(* IEC 61131-3 sources: kns-pump-station/tests/POUs/Station/FB_PumpRotation_Test, 30 files *)

(* ---- AdoptAtPlcStartFromFeedback.method.decl.st ---- *)
// 04 §13.3, PMI-35: старт ПЛК — подхват по ОС (GVL_IO.xP10n_RFB) до первого вызова устройства; запрос не снимается
// ни недоступностью первого цикла, ни ограничением последовательного пуска
METHOD PRIVATE AdoptAtPlcStartFromFeedback
VAR
    fbDut    : FB_PumpRotation;                    // ФБ под тестом
    fbTime   : PL.FB_FakeTime;                     // подменное время, старт 1 ч
    stCfg    : ST_StationCfg;                      // уставки по умолчанию (RunHours, tStagger 5 с)
    stRetain : ST_StationRetain;                   // следующий ведущий (Cyclic)
    afbPump  : ARRAY[1..3] OF FB_FakeMotorVfd;     // подменные насосы: доступны, Auto, готовы, стоят
    fbSink   : FB_FakeEventSink;                   // подменный журнал
END_VAR

(* ---- AdoptKeepsRunningPumpsOnAutoEntry.method.decl.st ---- *)
// 04 §3.2, PMI-30: вход в «Автомат» — роли получают работающие насосы (ещё в Manual в этом цикле), работающий не
// останавливается, ведущий — с меньшей наработкой
METHOD PRIVATE AdoptKeepsRunningPumpsOnAutoEntry
VAR
    fbDut    : FB_PumpRotation;                    // ФБ под тестом
    fbTime   : PL.FB_FakeTime;                     // подменное время, старт 1 ч
    stCfg    : ST_StationCfg;                      // уставки по умолчанию (RunHours, tStagger 5 с)
    stRetain : ST_StationRetain;                   // следующий ведущий (Cyclic)
    afbPump  : ARRAY[1..3] OF FB_FakeMotorVfd;     // подменные насосы: доступны, Auto, готовы, стоят
    fbSink   : FB_FakeEventSink;                   // подменный журнал
END_VAR

(* ---- Cycle.method.decl.st ---- *)
// Помощник: uiSteps шагов времени tStep с одним требуемым числом. xPlant — подменные насосы в Auto
// следуют запросам: работают, если запрошены, доступны и без отказа (видно со следующего шага)
METHOD PRIVATE Cycle
VAR_IN_OUT
    fbDut    : FB_PumpRotation;                 // ФБ под тестом
    fbTime   : PL.FB_FakeTime;                  // подменное время
    stCfg    : ST_StationCfg;                   // уставки
    stRetain : ST_StationRetain;                // энергонезависимые данные
    afbPump  : ARRAY[1..3] OF FB_FakeMotorVfd;  // подменные насосы
END_VAR
VAR_INPUT
    uiRequired : UINT;                          // требуемое число насосов
    tStep      : TIME;                          // шаг времени
    uiSteps    : UINT;                          // шагов
    xPlant     : BOOL;                          // насосы следуют запросам
END_VAR
VAR
    uiStep : UINT;                              // номер шага
    uiIdx  : UINT;                              // насос
END_VAR

(* ---- Cycle.method.impl.st ---- *)
FOR uiStep := 1 TO uiSteps DO
    fbTime.Advance(tStep := tStep);
    fbDut(uiRequired := uiRequired, itfTime := fbTime, stCfg := stCfg, stRetain := stRetain);
    IF xPlant THEN
        FOR uiIdx := 1 TO 3 DO
            IF afbPump[uiIdx].eMode = PL.E_DeviceMode.Auto THEN
                afbPump[uiIdx].xRunning := fbDut.axRun[uiIdx] AND afbPump[uiIdx].xAvailable
                                           AND NOT afbPump[uiIdx].xFault;
            END_IF
        END_FOR
    END_IF
END_FOR

(* ---- CyclicAdvancesNextLeadRetained.method.decl.st ---- *)
// 04 §8.1, PMI-10: по кругу — ведущий после stStationRetain.uiNextLead независимо от наработки, следующий
// запоминается энергонезависимо
METHOD PRIVATE CyclicAdvancesNextLeadRetained
VAR
    fbDut    : FB_PumpRotation;                    // ФБ под тестом
    fbTime   : PL.FB_FakeTime;                     // подменное время, старт 1 ч
    stCfg    : ST_StationCfg;                      // уставки по умолчанию (RunHours, tStagger 5 с)
    stRetain : ST_StationRetain;                   // следующий ведущий (Cyclic)
    afbPump  : ARRAY[1..3] OF FB_FakeMotorVfd;     // подменные насосы: доступны, Auto, готовы, стоят
    fbSink   : FB_FakeEventSink;                   // подменный журнал
END_VAR

(* ---- CyclicNextLeadFollowsRoleTransfer.method.decl.st ---- *)
// 04 §8.1, §8.2, PMI-10, PMI-11: по кругу следующий ведущий отсчитывается от насоса, который стал ведущим, в том
// числе без нового пуска (передача роли по ограничению непрерывной работы). Иначе после передачи Н1 → Н2
// следующий пуск снова достался бы Н2, а Н3 простаивал бы
METHOD PRIVATE CyclicNextLeadFollowsRoleTransfer
VAR
    fbDut    : FB_PumpRotation;                    // ФБ под тестом
    fbTime   : PL.FB_FakeTime;                     // подменное время, старт 1 ч
    stCfg    : ST_StationCfg;                      // уставки по умолчанию, режим Cyclic
    stRetain : ST_StationRetain;                   // следующий ведущий (Cyclic)
    afbPump  : ARRAY[1..3] OF FB_FakeMotorVfd;     // подменные насосы: доступны, Auto, готовы, стоят
    fbSink   : FB_FakeEventSink;                   // подменный журнал
END_VAR

(* ---- CyclicStopsAssist.method.decl.st ---- *)
// 04 §5.2: по кругу и без чередования — при уменьшении останавливается подпорный
METHOD PRIVATE CyclicStopsAssist
VAR
    fbDut    : FB_PumpRotation;                    // ФБ под тестом
    fbTime   : PL.FB_FakeTime;                     // подменное время, старт 1 ч
    stCfg    : ST_StationCfg;                      // уставки по умолчанию (RunHours, tStagger 5 с)
    stRetain : ST_StationRetain;                   // следующий ведущий (Cyclic)
    afbPump  : ARRAY[1..3] OF FB_FakeMotorVfd;     // подменные насосы: доступны, Auto, готовы, стоят
    fbSink   : FB_FakeEventSink;                   // подменный журнал
END_VAR

(* ---- DisabledNoRequestsRolesStandby.method.decl.st ---- *)
// DESIGN 6.5: станция не в «Автомате» — запросов нет, роли считаются (Standby у доступных, None у недоступных)
METHOD PRIVATE DisabledNoRequestsRolesStandby
VAR
    fbDut    : FB_PumpRotation;                    // ФБ под тестом
    fbTime   : PL.FB_FakeTime;                     // подменное время, старт 1 ч
    stCfg    : ST_StationCfg;                      // уставки по умолчанию (RunHours, tStagger 5 с)
    stRetain : ST_StationRetain;                   // следующий ведущий (Cyclic)
    afbPump  : ARRAY[1..3] OF FB_FakeMotorVfd;     // подменные насосы: доступны, Auto, готовы, стоят
    fbSink   : FB_FakeEventSink;                   // подменный журнал
END_VAR

(* ---- EmergencyRequiresAllThree.method.decl.st ---- *)
// 04 §10.2, PMI-20: аварийный режим — запросы всем трём насосам по одному через tStagger; роли Lead, Assist,
// Assist
METHOD PRIVATE EmergencyRequiresAllThree
VAR
    fbDut    : FB_PumpRotation;                    // ФБ под тестом
    fbTime   : PL.FB_FakeTime;                     // подменное время, старт 1 ч
    stCfg    : ST_StationCfg;                      // уставки по умолчанию (RunHours, tStagger 5 с)
    stRetain : ST_StationRetain;                   // следующий ведущий (Cyclic)
    afbPump  : ARRAY[1..3] OF FB_FakeMotorVfd;     // подменные насосы: доступны, Auto, готовы, стоят
    fbSink   : FB_FakeEventSink;                   // подменный журнал
END_VAR

(* ---- FaultedPumpLosesRequestImmediately.method.decl.st ---- *)
// 04 §9.1, PMI-12, PMI-13: отказавший ведущий теряет запрос сразу (роль None), замена — в том же вызове
METHOD PRIVATE FaultedPumpLosesRequestImmediately
VAR
    fbDut    : FB_PumpRotation;                    // ФБ под тестом
    fbTime   : PL.FB_FakeTime;                     // подменное время, старт 1 ч
    stCfg    : ST_StationCfg;                      // уставки по умолчанию (RunHours, tStagger 5 с)
    stRetain : ST_StationRetain;                   // следующий ведущий (Cyclic)
    afbPump  : ARRAY[1..3] OF FB_FakeMotorVfd;     // подменные насосы: доступны, Auto, готовы, стоят
    fbSink   : FB_FakeEventSink;                   // подменный журнал
END_VAR

(* ---- FixedOrder.method.decl.st ---- *)
// 04 §8.1: без чередования — Н1, Н2, Н3 по порядку; недоступный пропускается
METHOD PRIVATE FixedOrder
VAR
    fbDut    : FB_PumpRotation;                    // ФБ под тестом
    fbTime   : PL.FB_FakeTime;                     // подменное время, старт 1 ч
    stCfg    : ST_StationCfg;                      // уставки по умолчанию (RunHours, tStagger 5 с)
    stRetain : ST_StationRetain;                   // следующий ведущий (Cyclic)
    afbPump  : ARRAY[1..3] OF FB_FakeMotorVfd;     // подменные насосы: доступны, Auto, готовы, стоят
    fbSink   : FB_FakeEventSink;                   // подменный журнал
END_VAR

(* ---- ForeignRunningReducesRequests.method.decl.st ---- *)
// 04 §5.1, PMI-31: сторонний работающий насос (не в Auto) уменьшает число запросов станции
METHOD PRIVATE ForeignRunningReducesRequests
VAR
    fbDut    : FB_PumpRotation;                    // ФБ под тестом
    fbTime   : PL.FB_FakeTime;                     // подменное время, старт 1 ч
    stCfg    : ST_StationCfg;                      // уставки по умолчанию (RunHours, tStagger 5 с)
    stRetain : ST_StationRetain;                   // следующий ведущий (Cyclic)
    afbPump  : ARRAY[1..3] OF FB_FakeMotorVfd;     // подменные насосы: доступны, Auto, готовы, стоят
    fbSink   : FB_FakeEventSink;                   // подменный журнал
END_VAR

(* ---- GarbageNextLeadSanitized.method.decl.st ---- *)
// Мусор persistent-памяти: следующий ведущий вне 1…3 — с первого насоса
METHOD PRIVATE GarbageNextLeadSanitized
VAR
    fbDut    : FB_PumpRotation;                    // ФБ под тестом
    fbTime   : PL.FB_FakeTime;                     // подменное время, старт 1 ч
    stCfg    : ST_StationCfg;                      // уставки по умолчанию (RunHours, tStagger 5 с)
    stRetain : ST_StationRetain;                   // следующий ведущий (Cyclic)
    afbPump  : ARRAY[1..3] OF FB_FakeMotorVfd;     // подменные насосы: доступны, Auto, готовы, стоят
    fbSink   : FB_FakeEventSink;                   // подменный журнал
END_VAR

(* ---- HandoverAfterTMaxContRunWithOverlap.method.decl.st ---- *)
// 04 §8.2, PMI-11: ведущий работает непрерывно tMaxContRun — пускается резервный, через tOverlap после его ОС
// прежний останавливается, роль у замены; событие 101007
METHOD PRIVATE HandoverAfterTMaxContRunWithOverlap
VAR
    fbDut    : FB_PumpRotation;                    // ФБ под тестом
    fbTime   : PL.FB_FakeTime;                     // подменное время, старт 1 ч
    stCfg    : ST_StationCfg;                      // уставки по умолчанию (RunHours, tStagger 5 с)
    stRetain : ST_StationRetain;                   // следующий ведущий (Cyclic)
    afbPump  : ARRAY[1..3] OF FB_FakeMotorVfd;     // подменные насосы: доступны, Auto, готовы, стоят
    fbSink   : FB_FakeEventSink;                   // подменный журнал
END_VAR

(* ---- HandoverDisabledInEmergency.method.decl.st ---- *)
// 04 §8.2: передача роли не выполняется в аварийном режиме, по поплавкам и при последовательном пуске
// (xHandoverAllowed = FALSE); tMaxContRun = 0 — выключено
METHOD PRIVATE HandoverDisabledInEmergency
VAR
    fbDut    : FB_PumpRotation;                    // ФБ под тестом
    fbTime   : PL.FB_FakeTime;                     // подменное время, старт 1 ч
    stCfg    : ST_StationCfg;                      // уставки по умолчанию (RunHours, tStagger 5 с)
    stRetain : ST_StationRetain;                   // следующий ведущий (Cyclic)
    afbPump  : ARRAY[1..3] OF FB_FakeMotorVfd;     // подменные насосы: доступны, Auto, готовы, стоят
    fbSink   : FB_FakeEventSink;                   // подменный журнал
    fbDut2   : FB_PumpRotation;                    // второй экземпляр: tMaxContRun = 0
    stCfg0   : ST_StationCfg;                      // уставки с tMaxContRun = 0
END_VAR

(* ---- HandoverLeadNeedsCommInPid.method.decl.st ---- *)
// 04 §5.2 п. 3, §8.2, §12, PMI-11: в ПИД замена ведущего при передаче роли — только готовый насос со связью с ПЧ.
// Резерв без связи роль не получает (иначе после перекрытия ведущим стал бы насос без связи, ПИД потерял бы
// готовность и станция ушла бы в ступенчатое с KNS1.STEP) — повтор через STN_HANDOVER_RETRY
METHOD PRIVATE HandoverLeadNeedsCommInPid
VAR
    fbDut    : FB_PumpRotation;                    // ФБ под тестом
    fbTime   : PL.FB_FakeTime;                     // подменное время, старт 1 ч
    stCfg    : ST_StationCfg;                      // уставки по умолчанию (RunHours, tStagger 5 с)
    stRetain : ST_StationRetain;                   // следующий ведущий (Cyclic)
    afbPump  : ARRAY[1..3] OF FB_FakeMotorVfd;     // подменные насосы: доступны, Auto, готовы, стоят
    fbSink   : FB_FakeEventSink;                   // подменный журнал
END_VAR

(* ---- HandoverRetryWhenNoStandby.method.decl.st ---- *)
// 04 §8.2: резерва нет — длительно работавший продолжает, повтор через STN_HANDOVER_RETRY = 10 мин, не раньше
METHOD PRIVATE HandoverRetryWhenNoStandby
VAR
    fbDut    : FB_PumpRotation;                    // ФБ под тестом
    fbTime   : PL.FB_FakeTime;                     // подменное время, старт 1 ч
    stCfg    : ST_StationCfg;                      // уставки по умолчанию (RunHours, tStagger 5 с)
    stRetain : ST_StationRetain;                   // следующий ведущий (Cyclic)
    afbPump  : ARRAY[1..3] OF FB_FakeMotorVfd;     // подменные насосы: доступны, Auto, готовы, стоят
    fbSink   : FB_FakeEventSink;                   // подменный журнал
END_VAR

(* ---- LeadSwapWithoutStartStop.method.decl.st ---- *)
// 04 §12, PMI-28: у ведущего пропала связь, у работающего подпорного она есть — смена ведущего без пуска и
// останова (101005)
METHOD PRIVATE LeadSwapWithoutStartStop
VAR
    fbDut    : FB_PumpRotation;                    // ФБ под тестом
    fbTime   : PL.FB_FakeTime;                     // подменное время, старт 1 ч
    stCfg    : ST_StationCfg;                      // уставки по умолчанию (RunHours, tStagger 5 с)
    stRetain : ST_StationRetain;                   // следующий ведущий (Cyclic)
    afbPump  : ARRAY[1..3] OF FB_FakeMotorVfd;     // подменные насосы: доступны, Auto, готовы, стоят
    fbSink   : FB_FakeEventSink;                   // подменный журнал
END_VAR

(* ---- ReadyBeforeInhibited.method.decl.st ---- *)
// 04 §5.2: сначала готовые к пуску, затем доступные в паузе (запрос подождёт)
METHOD PRIVATE ReadyBeforeInhibited
VAR
    fbDut    : FB_PumpRotation;                    // ФБ под тестом
    fbTime   : PL.FB_FakeTime;                     // подменное время, старт 1 ч
    stCfg    : ST_StationCfg;                      // уставки по умолчанию (RunHours, tStagger 5 с)
    stRetain : ST_StationRetain;                   // следующий ведущий (Cyclic)
    afbPump  : ARRAY[1..3] OF FB_FakeMotorVfd;     // подменные насосы: доступны, Auto, готовы, стоят
    fbSink   : FB_FakeEventSink;                   // подменный журнал
END_VAR

(* ---- RequestLimitCapsRequests.method.decl.st ---- *)
// 04 §13.2, PMI-34: последовательный пуск — новых запросов не больше uiRequestLimit
METHOD PRIVATE RequestLimitCapsRequests
VAR
    fbDut    : FB_PumpRotation;                    // ФБ под тестом
    fbTime   : PL.FB_FakeTime;                     // подменное время, старт 1 ч
    stCfg    : ST_StationCfg;                      // уставки по умолчанию (RunHours, tStagger 5 с)
    stRetain : ST_StationRetain;                   // следующий ведущий (Cyclic)
    afbPump  : ARRAY[1..3] OF FB_FakeMotorVfd;     // подменные насосы: доступны, Auto, готовы, стоят
    fbSink   : FB_FakeEventSink;                   // подменный журнал
END_VAR

(* ---- RequireCommPicksCommPumpAsLead.method.decl.st ---- *)
// 04 §5.2, §12, PMI-28: в ПИД ведущим назначается насос со связью с ПЧ, даже если у насоса без связи наработка
// меньше
METHOD PRIVATE RequireCommPicksCommPumpAsLead
VAR
    fbDut    : FB_PumpRotation;                    // ФБ под тестом
    fbTime   : PL.FB_FakeTime;                     // подменное время, старт 1 ч
    stCfg    : ST_StationCfg;                      // уставки по умолчанию (RunHours, tStagger 5 с)
    stRetain : ST_StationRetain;                   // следующий ведущий (Cyclic)
    afbPump  : ARRAY[1..3] OF FB_FakeMotorVfd;     // подменные насосы: доступны, Auto, готовы, стоят
    fbSink   : FB_FakeEventSink;                   // подменный журнал
END_VAR

(* ---- ResetPumpBecomesStandby.method.decl.st ---- *)
// 04 §9.1, PMI-12: после сброса отказа насос резервный и сам не пускается
METHOD PRIVATE ResetPumpBecomesStandby
VAR
    fbDut    : FB_PumpRotation;                    // ФБ под тестом
    fbTime   : PL.FB_FakeTime;                     // подменное время, старт 1 ч
    stCfg    : ST_StationCfg;                      // уставки по умолчанию (RunHours, tStagger 5 с)
    stRetain : ST_StationRetain;                   // следующий ведущий (Cyclic)
    afbPump  : ARRAY[1..3] OF FB_FakeMotorVfd;     // подменные насосы: доступны, Auto, готовы, стоят
    fbSink   : FB_FakeEventSink;                   // подменный журнал
END_VAR

(* ---- RunHoursPicksLeastHours.method.decl.st ---- *)
// 04 §8.1, PMI-09: чередование по моточасам — ведущим при пуске назначается насос с наименьшей наработкой; событие
// 101005 с его номером
METHOD PRIVATE RunHoursPicksLeastHours
VAR
    fbDut    : FB_PumpRotation;                    // ФБ под тестом
    fbTime   : PL.FB_FakeTime;                     // подменное время, старт 1 ч
    stCfg    : ST_StationCfg;                      // уставки по умолчанию (RunHours, tStagger 5 с)
    stRetain : ST_StationRetain;                   // следующий ведущий (Cyclic)
    afbPump  : ARRAY[1..3] OF FB_FakeMotorVfd;     // подменные насосы: доступны, Auto, готовы, стоят
    fbSink   : FB_FakeEventSink;                   // подменный журнал
END_VAR

(* ---- RunningKeepRoles.method.decl.st ---- *)
// 04 §5.2: роли работающих по запросу насосов сохраняются, даже если наработка другого стала меньше
METHOD PRIVATE RunningKeepRoles
VAR
    fbDut    : FB_PumpRotation;                    // ФБ под тестом
    fbTime   : PL.FB_FakeTime;                     // подменное время, старт 1 ч
    stCfg    : ST_StationCfg;                      // уставки по умолчанию (RunHours, tStagger 5 с)
    stRetain : ST_StationRetain;                   // следующий ведущий (Cyclic)
    afbPump  : ARRAY[1..3] OF FB_FakeMotorVfd;     // подменные насосы: доступны, Auto, готовы, стоят
    fbSink   : FB_FakeEventSink;                   // подменный журнал
END_VAR

(* ---- StaggerDelaysSecondStart.method.decl.st ---- *)
// 04 §5.2: несколько пусков — по одному с интервалом tStagger = 5 с (ровно на 5 с, не раньше); xStaggerWait во
// время ожидания
METHOD PRIVATE StaggerDelaysSecondStart
VAR
    fbDut    : FB_PumpRotation;                    // ФБ под тестом
    fbTime   : PL.FB_FakeTime;                     // подменное время, старт 1 ч
    stCfg    : ST_StationCfg;                      // уставки по умолчанию (RunHours, tStagger 5 с)
    stRetain : ST_StationRetain;                   // следующий ведущий (Cyclic)
    afbPump  : ARRAY[1..3] OF FB_FakeMotorVfd;     // подменные насосы: доступны, Auto, готовы, стоят
    fbSink   : FB_FakeEventSink;                   // подменный журнал
END_VAR

(* ---- StaggerSkippedWhenPreviousDropped.method.decl.st ---- *)
// 04 §5.2, §9.1: насос предыдущего нового запроса отказал при пуске — замена без ожидания tStagger
METHOD PRIVATE StaggerSkippedWhenPreviousDropped
VAR
    fbDut    : FB_PumpRotation;                    // ФБ под тестом
    fbTime   : PL.FB_FakeTime;                     // подменное время, старт 1 ч
    stCfg    : ST_StationCfg;                      // уставки по умолчанию (RunHours, tStagger 5 с)
    stRetain : ST_StationRetain;                   // следующий ведущий (Cyclic)
    afbPump  : ARRAY[1..3] OF FB_FakeMotorVfd;     // подменные насосы: доступны, Auto, готовы, стоят
    fbSink   : FB_FakeEventSink;                   // подменный журнал
END_VAR

(* ---- StopKeepsCommPumpInPid.method.decl.st ---- *)
// 04 §5.2 п. 3, §12, PMI-05, PMI-28: в ПИД при снятии роли по моточасам насос со связью с ПЧ снимается последним.
// Иначе остался бы насос без связи: ПИД потерял бы готовность и станция ушла бы в ступенчатое с KNS1.STEP, хотя
// работал насос со связью
METHOD PRIVATE StopKeepsCommPumpInPid
VAR
    fbDut    : FB_PumpRotation;                    // ФБ под тестом
    fbTime   : PL.FB_FakeTime;                     // подменное время, старт 1 ч
    stCfg    : ST_StationCfg;                      // уставки по умолчанию (RunHours, tStagger 5 с)
    stRetain : ST_StationRetain;                   // следующий ведущий (Cyclic)
    afbPump  : ARRAY[1..3] OF FB_FakeMotorVfd;     // подменные насосы: доступны, Auto, готовы, стоят
    fbSink   : FB_FakeEventSink;                   // подменный журнал
END_VAR

(* ---- StopMoreHoursWhenFewerNeeded.method.decl.st ---- *)
// 04 §5.2, PMI-03: нужно меньше насосов — останавливается насос с большей наработкой; если это ведущий, роль
// переходит к оставшемуся (101005)
METHOD PRIVATE StopMoreHoursWhenFewerNeeded
VAR
    fbDut    : FB_PumpRotation;                    // ФБ под тестом
    fbTime   : PL.FB_FakeTime;                     // подменное время, старт 1 ч
    stCfg    : ST_StationCfg;                      // уставки по умолчанию (RunHours, tStagger 5 с)
    stRetain : ST_StationRetain;                   // следующий ведущий (Cyclic)
    afbPump  : ARRAY[1..3] OF FB_FakeMotorVfd;     // подменные насосы: доступны, Auto, готовы, стоят
    fbSink   : FB_FakeEventSink;                   // подменный журнал
END_VAR

(* ---- TieBreakStartsThenIndex.method.decl.st ---- *)
// 04 §8.1: при равной наработке — меньше пусков, при равных пусках — меньший номер
METHOD PRIVATE TieBreakStartsThenIndex
VAR
    fbDut    : FB_PumpRotation;                    // ФБ под тестом
    fbTime   : PL.FB_FakeTime;                     // подменное время, старт 1 ч
    stCfg    : ST_StationCfg;                      // уставки по умолчанию (RunHours, tStagger 5 с)
    stRetain : ST_StationRetain;                   // следующий ведущий (Cyclic)
    afbPump  : ARRAY[1..3] OF FB_FakeMotorVfd;     // подменные насосы: доступны, Auto, готовы, стоят
    fbSink   : FB_FakeEventSink;                   // подменный журнал
END_VAR

(* ---- TimeBackwardsRestartsStagger.method.decl.st ---- *)
// Время назад — интервал tStagger отсчитывается заново: два пуска подряд не выдаются
METHOD PRIVATE TimeBackwardsRestartsStagger
VAR
    fbDut    : FB_PumpRotation;                    // ФБ под тестом
    fbTime   : PL.FB_FakeTime;                     // подменное время, старт 1 ч
    stCfg    : ST_StationCfg;                      // уставки по умолчанию (RunHours, tStagger 5 с)
    stRetain : ST_StationRetain;                   // следующий ведущий (Cyclic)
    afbPump  : ARRAY[1..3] OF FB_FakeMotorVfd;     // подменные насосы: доступны, Auto, готовы, стоят
    fbSink   : FB_FakeEventSink;                   // подменный журнал
END_VAR
